(* IEC 61131-3 sources: volt/packages/volt-lsp-iec/test-corpus/lenze-mid/Device/Plc Logic/Application/Library Manager/CAA Device Diagnosis, 56 files *)

(* ---- BUS_INFO.dut ---- *)
TYPE BUS_INFO :
STRUCT
	ETYPE : BUS_TYPE;
	IDSYSTEM : CAA.IDENT;
	IDINSTANCE : CAA.IDENT;
END_STRUCT
END_TYPE

(* ---- BUS_STATE.dut ---- *)
TYPE BUS_STATE :
(
	UNKNOWN,
	STOPPED,
	RUNNING,
	ERROR,
	DISABLED
);
END_TYPE

(* ---- BUS_TYPE.dut ---- *)
TYPE BUS_TYPE :
(
	UNKNOWN := 16#0,
	PROFIBUS_DP := 16#1,
	CAN := 16#2,
	CANOPEN := 16#3,
	DEVICENET := 16#4,
	ETHERCAT := 16#5,
	PROFINET_IO := 16#6,
	ETHERNET_IP := 16#7,
	SERCOSII := 16#8,
	SERCOSIII := 16#9,
	MODBUS_TCP := 16#A,
	MODBUS_RTU := 16#B,
	AS_INTERFACE := 16#C,
	INTERBUS := 16#D,
	J1939 := 16#E,
	LON := 16#F,
	CC_LINK := 16#10,
	POWERLINK := 16#11,
	ETHERNET := 16#12,
	SERIAL_LINE := 16#13,
	VEN_SPEC := 16#14,
	FIRST_MF := 16#8000,
	LAST := 16#FFFF
);
END_TYPE

(* ---- DED_PNS_SUBMODULE_CFG.dut ---- *)
TYPE DED_PNS_SUBMODULE_CFG :
STRUCT
	UISLOT : UINT;
	UISUBSLOT : UINT;
	ULMODULEID : UDINT;
	ULSUBMODULEID : UDINT;
	ULPROVDATALEN : UDINT;
	ULCONSDATALEN : UDINT;
END_STRUCT
END_TYPE

(* ---- DEVICE_INFO.dut ---- *)
TYPE DEVICE_INFO :
STRUCT
	ETYPE : DEVICE_TYPE;
	IDSYSTEM : CAA.IDENT;
	IDINSTANCE : CAA.IDENT;
END_STRUCT
END_TYPE

(* ---- DEVICE_STATE.dut ---- *)
TYPE DEVICE_STATE :
(
	UNKNOWN,
	STOPPED,
	RUNNING,
	ERROR,
	DISABLED,
	NOT_CONFIGURED,
	CONFIGURED,
	NOT_FOUND
);
END_TYPE

(* ---- DEVICE_TRANSITION_STATE.dut ---- *)
TYPE DEVICE_TRANSITION_STATE :
(
	START,
	STOP,
	RESET
);
END_TYPE

(* ---- DEVICE_TYPE.dut ---- *)
TYPE DEVICE_TYPE :
(
	UNKNOWN := 16#0,
	FIELDBUS_MASTER := 16#1,
	FIELDBUS_SLAVE := 16#2,
	SAFETY_DEVICE := 16#3,
	SM_DEVICE := 16#4,
	SOFT_VISION_DEVICE := 16#5,
	DTM_DEVICE := 16#6,
	SPEC_IO_MODULE := 16#7,
	PLC := 16#1000,
	SAFETY_PLC := 16#1002,
	DRIVE := 16#1003,
	PARAM_DEVICE := 16#1004,
	HMI := 16#1005,
	SM_PLC := 16#1006
);
END_TYPE

(* ---- ERROR.dut ---- *)
TYPE ERROR :
(
	NO_ERROR := 0,
	FIRST_ERROR := 1300,
	TIME_OUT := 1301,
	ABORT := 1302,
	REF_INVALID := 1303,
	NOT_SUPPORTED := 1304,
	ERROR_IO := 1305,
	PARAM_INVALID := 1306,
	NODE_NOT_EXISTING := 1307,
	NO_MEMORY := 1308,
	ADR_NOT_FOUND := 1309,
	INST_NOT_FOUND := 1310,
	NO_DATA := 1311,
	OPERATION_INVALID := 1312,
	FIRST_MF := 1350,
	LAST_ERROR := 1399
);
END_TYPE

(* ---- ERROR_INFO.dut ---- *)
TYPE ERROR_INFO :
STRUCT
	IDERRORCODE : CAA.IDENT;
END_STRUCT
END_TYPE

(* ---- LOG_ENTRY.dut ---- *)
TYPE LOG_ENTRY :
STRUCT
	TKTIMESTAMP : CAA.TICK;
	IDMESSAGE : CAA.IDENT;
	IDSOURCE : CAA.IDENT;
END_STRUCT
END_TYPE

(* ---- LOGGER_MODE.dut ---- *)
TYPE LOGGER_MODE :
(
	LINEAR,
	CIRCULAR
);
END_TYPE

(* ---- PROC_CMD.dut ---- *)
TYPE PROC_CMD :
(
	NONE := 0,
	EXECUTE,
	ABORT
);
END_TYPE

(* ---- PROC_STATE.dut ---- *)
TYPE PROC_STATE :
(
	DORMAND := 0,
	BUSY,
	DONE,
	ABORTED,
	ERROR
);
END_TYPE

(* ---- QOS_INFO.dut ---- *)
TYPE QOS_INFO :
STRUCT
	CTERROR : CAA.COUNT;
	USIBUSLOAD : USINT;
END_STRUCT
END_TYPE

(* ---- TIDENTIFICATIONPARAMETER.dut ---- *)
TYPE TIDENTIFICATIONPARAMETER :
STRUCT
	IPADDRESS : ARRAY [0..3] OF BYTE;
	SUBNETMASK : ARRAY [0..3] OF BYTE;
	DEFAULTGATEWAY : ARRAY [0..3] OF BYTE;
	MACADDRESS : ARRAY [0..5] OF BYTE;
	STATIONNAME : STRING;
END_STRUCT
END_TYPE

(* ---- TISOCHRONEMODE.dut ---- *)
TYPE TISOCHRONEMODE :
STRUCT
	T_DC_BASE : UINT;
	T_DC_MIN : UINT;
	T_DC_MAX : UINT;
	T_IO_BASE : UDINT;
	T_IO_INPUTMIN : UDINT;
	T_IO_OUTPUTMIN : UDINT;
	ISOCHRONEMODEREQUIRED : BOOL;
END_STRUCT
END_TYPE

(* ---- TMODULEPARAMETER.dut ---- *)
TYPE TMODULEPARAMETER :
STRUCT
	MODULEIDENTNUMBER : UDINT;
	SLOTNUMBER : UINT;
	UINUMBERSUBMODULES : UINT;
END_STRUCT
END_TYPE

(* ---- TSLAVEPARAMETER.dut ---- *)
TYPE TSLAVEPARAMETER :
STRUCT
	UIDEVICEID : UINT;
	UIVENDORID : UINT;
	IDENTIFICATION : TIdentificationParameter;
	RTCLASS : UINT;
	VLANID : UINT;
	VLANPRIORITY : UINT;
	SENDCLOCK : UINT;
	REDUCTIONRATIO : UINT;
	WATCHDOGINTERVAL : UINT;
	MULTIPLEWRITESUPPORTED : BOOL;
	IOXSREQUIRED : BOOL;
	MAXINPUTLENGTH : UINT;
	MAXOUTPUTLENGTH : UINT;
	MAXDATALENGTH : UINT;
	UIMINSLAVEINTERVAL : UINT;
	UIOBJECTUUIDINSTANCE : UINT;
END_STRUCT
END_TYPE

(* ---- TVIRTUALSUBMODULE.dut ---- *)
TYPE TVIRTUALSUBMODULE :
STRUCT
	SUBMODULEIDENTNUMBER : UDINT;
	SUBSLOTNUMBER : UINT;
	API : UDINT;
	PROFISAFESUPPORTED : BOOL;
	ISOCHRONEMODE : TIsochroneMode;
	UINUMBERRDI : UINT;
	UISUBMODULEPROP : UINT;
	USIIOPSLEN : USINT;
	USIIOCSLEN : USINT;
END_STRUCT
END_TYPE

(* ---- DEVICEDIAGNOSISGLOBALS.gvl ---- *)
VAR_GLOBAL
	G_ITFROOTINODEINST : POINTER TO INode;
	G_ITFROOTNODECOUNT : UDINT;
END_VAR

(* ---- ERROR_CODES.gvl ---- *)
VAR_GLOBAL
	EC_NO_ERROR : CAA.IDENT := 16#0;
	EC_FIRST_INFO : CAA.IDENT := 16#1000;
	EC_LAST_INFO : CAA.IDENT := 16#1FFF;
	EC_FIRST_WARNING : CAA.IDENT := 16#2000;
	EC_LAST_WARNING : CAA.IDENT := 16#2FFF;
	EC_FIRST_ERROR : CAA.IDENT := 16#3000;
	EC_LAST_ERROR : CAA.IDENT := 16#3FFF;
	EC_FIRST_EMCY : CAA.IDENT := 16#4000;
	EC_LAST_EMCY : CAA.IDENT := 16#4FFF;
END_VAR

(* ---- VERSIONCONSTANTS.gvl ---- *)
VAR_GLOBAL
	GC_BYVERSION : BYTE := 1;
	GC_BYVERSION_1 : BYTE := 1;
END_VAR

(* ---- IBUS.itf ---- *)
INTERFACE IBUS
END_INTERFACE

METHOD GETBUSDIAGNOSISINFO : ERROR
VAR_INPUT
	PDATA : CAA.PVOID;
	SZSIZE : CAA.SIZE;
END_VAR
VAR_OUTPUT
	SZCOUNT : CAA.SIZE;
END_VAR
END_METHOD

METHOD GETBUSERRORASYNC : PROC_STATE
VAR_INPUT
	ECMD : PROC_CMD;
END_VAR
VAR_OUTPUT
	EERROR : ERROR;
END_VAR
VAR_IN_OUT
	ERIBUSERROR : ERROR_INFO;
END_VAR
END_METHOD

METHOD GETBUSINFO : ERROR
VAR_IN_OUT
	BUIINFO : BUS_INFO;
END_VAR
END_METHOD

METHOD GETBUSSTATE : BUS_STATE
VAR_OUTPUT
	XDIAGNOSISINFOAVAILABLE : BOOL;
	EERROR : ERROR;
END_VAR
END_METHOD

METHOD GETQOS : ERROR
VAR_IN_OUT
	QUALITYINFO : QOS_INFO;
END_VAR
END_METHOD

METHOD GETSPECIFICBUSSTATE : ERROR
VAR_INPUT
	PDATA : CAA.PVOID;
	SZSIZE : CAA.SIZE;
END_VAR
VAR_OUTPUT
	SZCOUNT : CAA.SIZE;
END_VAR
END_METHOD

(* ---- IDEVICE.itf ---- *)
INTERFACE IDEVICE
END_INTERFACE

METHOD GETDEVICEDIAGNOSISINFO : ERROR
VAR_INPUT
	PDATA : CAA.PVOID;
	SZSIZE : CAA.SIZE;
END_VAR
VAR_OUTPUT
	SZCOUNT : CAA.SIZE;
END_VAR
END_METHOD

METHOD GETDEVICEERRORASYNC : PROC_STATE
VAR_INPUT
	ECMD : PROC_CMD;
END_VAR
VAR_OUTPUT
	EERROR : ERROR;
END_VAR
VAR_IN_OUT
	ERIDEVICEERROR : ERROR_INFO;
END_VAR
END_METHOD

METHOD GETDEVICEINFO : ERROR
VAR_IN_OUT
	DEIINFO : DEVICE_INFO;
END_VAR
END_METHOD

METHOD GETDEVICESTATE : DEVICE_STATE
VAR_OUTPUT
	XDIAGNOSISINFOAVAILABLE : BOOL;
	EERROR : ERROR;
END_VAR
END_METHOD

METHOD SETCOMMUNICATIONSTATE : ERROR
VAR_INPUT
	EREQUESTEDSTATE : DEVICE_TRANSITION_STATE;
END_VAR
END_METHOD

METHOD GETSPECIFICDEVICEERRORASYNC : PROC_STATE
VAR_INPUT
	ECMD : PROC_CMD;
	PDATA : CAA.PVOID;
	SZSIZE : CAA.SIZE;
END_VAR
VAR_OUTPUT
	SZCOUNT : CAA.SIZE;
	EERROR : ERROR;
END_VAR
END_METHOD

METHOD GETSPECIFICDEVICESTATE : ERROR
VAR_INPUT
	PDATA : CAA.PVOID;
	SZSIZE : CAA.SIZE;
END_VAR
VAR_OUTPUT
	SZCOUNT : CAA.SIZE;
END_VAR
END_METHOD

(* ---- IDEVICE2.itf ---- *)
INTERFACE IDEVICE2
END_INTERFACE

METHOD CHECKCURRENTSUPPORTEDCOMMUNICATIONSTATE : BOOL
VAR_INPUT
	EREQUESTEDSTATE : DEVICE_TRANSITION_STATE;
END_VAR
END_METHOD

METHOD CHECKSUPPORTEDCOMMUNICATIONSTATE : BOOL
VAR_INPUT
	EREQUESTEDSTATE : DEVICE_TRANSITION_STATE;
END_VAR
END_METHOD

(* ---- ILOGGER.itf ---- *)
INTERFACE ILOGGER
END_INTERFACE

METHOD DISABLELOGGER : ERROR
END_METHOD

METHOD ENABLELOGGER : ERROR
VAR_INPUT
	EMODE : LOGGER_MODE;
	CTMAXLOGMESSAGES : CAA.COUNT;
END_VAR
END_METHOD

METHOD GETLOGENTRY : ERROR
VAR_IN_OUT
	LOGENTRY : LOG_ENTRY;
END_VAR
END_METHOD

(* ---- INODE.itf ---- *)
INTERFACE INODE
END_INTERFACE

METHOD GETCHILD : INode
VAR_INPUT
	UDIINDEX : UDINT;
END_VAR
END_METHOD

METHOD INITIALIZE_DIAG : UDINT
VAR_INPUT
	PCONNECTOR : POINTER TO IoConfigConnector;
	NCONNECTORCOUNT : DINT;
	PARENT : POINTER TO INode;
	CHILDREN : POINTER TO INode;
	UDICHILDCOUNT : UDINT;
END_VAR
END_METHOD

(* ---- IRECONFIGUREPROVIDER.itf ---- *)
INTERFACE IRECONFIGUREPROVIDER
END_INTERFACE

METHOD RECONFIGUREASYNC : PROC_STATE
VAR_INPUT
	ECMD : PROC_CMD;
	ITFSENDER : INode;
END_VAR
VAR_OUTPUT
	EERROR : ERROR;
END_VAR
END_METHOD

METHOD REGISTERIRPCHILD : ERROR
VAR_INPUT
	ITFCHILD : IReconfigureProvider;
END_VAR
END_METHOD

(* ---- ISTACK.itf ---- *)
INTERFACE ISTACK
END_INTERFACE

METHOD GETBUSSCANASYNC : PROC_STATE
VAR_INPUT
	ECMD : PROC_CMD;
END_VAR
VAR_OUTPUT
	ITFFIRSTDEVICE : INode;
	EERROR : ERROR;
END_VAR
END_METHOD

METHOD GETLOGGER : ILogger
VAR_OUTPUT
	EERROR : ERROR;
END_VAR
END_METHOD

(* ---- CANRECONFIGURE.pou ---- *)
FUNCTION CANRECONFIGURE : BOOL
VAR_INPUT
	ITFNODE : INode;
END_VAR
END_FUNCTION

(* ---- GETDEVICENAMESTRING.pou ---- *)
FUNCTION GETDEVICENAMESTRING : STRING
VAR_INPUT
	ITFNODE : INode;
END_VAR
END_FUNCTION

(* ---- GETDEVICENAMEWSTRING.pou ---- *)
FUNCTION GETDEVICENAMEWSTRING : WSTRING
VAR_INPUT
	ITFNODE : INode;
END_VAR
END_FUNCTION

(* ---- GETNEXTNODE.pou ---- *)
FUNCTION GETNEXTNODE : INode
VAR_INPUT
	ITFCURRENT : INode;
END_VAR
END_FUNCTION

(* ---- GETNODEDEPTH.pou ---- *)
FUNCTION GETNODEDEPTH : INT
VAR_INPUT
	ITFNODE : INode;
END_VAR
END_FUNCTION

(* ---- GETROOT.pou ---- *)
FUNCTION GETROOT : INode
END_FUNCTION

(* ---- GETSUPPLIERVERSION.pou ---- *)
FUNCTION GETSUPPLIERVERSION : WORD
VAR_INPUT
	XDUMMY : BOOL;
END_VAR
END_FUNCTION

(* ---- INODE_TO_IBUS.pou ---- *)
FUNCTION INODE_TO_IBUS : IBus
VAR_INPUT
	ITFNODE : INode;
END_VAR
END_FUNCTION

(* ---- INODE_TO_IDEVICE.pou ---- *)
FUNCTION INODE_TO_IDEVICE : IDevice
VAR_INPUT
	ITFNODE : INode;
END_VAR
END_FUNCTION

(* ---- INODE_TO_IDEVICE2.pou ---- *)
FUNCTION INODE_TO_IDEVICE2 : IDevice2
VAR_INPUT
	ITFNODE : INode;
END_VAR
END_FUNCTION

(* ---- INODE_TO_ISTACK.pou ---- *)
FUNCTION INODE_TO_ISTACK : IStack
VAR_INPUT
	ITFNODE : INode;
END_VAR
END_FUNCTION

(* ---- ISCONNECTORENABLED.pou ---- *)
FUNCTION ISCONNECTORENABLED : BOOL
VAR_INPUT
	PCONNECTOR : POINTER TO IoStandard.IoConfigConnector;
END_VAR
END_FUNCTION

(* ---- CAADIAGDEVICEDEFAULT.pou ---- *)
FUNCTION_BLOCK CAADIAGDEVICEDEFAULT EXTENDS CAADiagTreeBase
VAR
	M_DIAG : CAADiagnosisBase;
	_DEIINFO : DEVICE_INFO;
END_VAR
END_FUNCTION_BLOCK

METHOD CHECKCURRENTSUPPORTEDCOMMUNICATIONSTATE : BOOL
VAR_INPUT
	EREQUESTEDSTATE : DEVICE_TRANSITION_STATE;
END_VAR
END_METHOD

METHOD CHECKSUPPORTEDCOMMUNICATIONSTATE : BOOL
VAR_INPUT
	EREQUESTEDSTATE : DEVICE_TRANSITION_STATE;
END_VAR
END_METHOD

METHOD GETDEVICEDIAGNOSISINFO : ERROR
VAR_INPUT
	PDATA : CAA.PVOID;
	SZSIZE : CAA.SIZE;
END_VAR
VAR_OUTPUT
	SZCOUNT : CAA.SIZE;
END_VAR
END_METHOD

METHOD GETDEVICEERRORASYNC : PROC_STATE
VAR_INPUT
	ECMD : PROC_CMD;
END_VAR
VAR_OUTPUT
	EERROR : ERROR;
END_VAR
VAR_IN_OUT
	ERIDEVICEERROR : ERROR_INFO;
END_VAR
END_METHOD

METHOD GETDEVICEINFO : ERROR
VAR_IN_OUT
	DEIINFO : DEVICE_INFO;
END_VAR
END_METHOD

METHOD GETDEVICESTATE : DEVICE_STATE
VAR_OUTPUT
	XDIAGNOSISINFOAVAILABLE : BOOL;
	EERROR : ERROR;
END_VAR
END_METHOD

METHOD GETPROFINETDEVICEINFO : ERROR
VAR_IN_OUT
	DEIINFO : DEVICE_INFO;
END_VAR
END_METHOD

METHOD GETSPECIFICDEVICEERRORASYNC : PROC_STATE
VAR_INPUT
	ECMD : PROC_CMD;
	PDATA : CAA.PVOID;
	SZSIZE : CAA.SIZE;
END_VAR
VAR_OUTPUT
	SZCOUNT : CAA.SIZE;
	EERROR : ERROR;
END_VAR
END_METHOD

METHOD GETSPECIFICDEVICESTATE : ERROR
VAR_INPUT
	PDATA : CAA.PVOID;
	SZSIZE : CAA.SIZE;
END_VAR
VAR_OUTPUT
	SZCOUNT : CAA.SIZE;
END_VAR
END_METHOD

METHOD INITIALIZE_DIAG : UDINT
VAR_INPUT
	PCONNECTOR : POINTER TO IoConfigConnector;
	NCONNECTORCOUNT : DINT;
	PARENT : POINTER TO INode;
	CHILDREN : POINTER TO INode;
	UDICHILDCOUNT : UDINT;
END_VAR
END_METHOD

METHOD SETCOMMUNICATIONSTATE : ERROR
VAR_INPUT
	EREQUESTEDSTATE : DEVICE_TRANSITION_STATE;
END_VAR
END_METHOD

(* ---- CAADIAGNOSISBASE.pou ---- *)
FUNCTION_BLOCK CAADIAGNOSISBASE
VAR
	M_NCOUNT : DINT;
	M_PCONNECTOR : POINTER TO IoConfigConnector;
	BUSLOGGER : Logger;
END_VAR
END_FUNCTION_BLOCK

METHOD CALCIPADRUDINT : UDINT
VAR_INPUT
	PABY : POINTER TO ARRAY [0..3] OF BYTE;
END_VAR
END_METHOD

METHOD GETBUSINFO : ERROR
VAR_IN_OUT
	BUIINFO : BUS_INFO;
END_VAR
END_METHOD

METHOD GETBUSSCANASYNC : PROC_STATE
VAR_INPUT
	ECMD : PROC_CMD;
END_VAR
VAR_OUTPUT
	ITFFIRSTDEVICE : INode;
	EERROR : ERROR;
END_VAR
END_METHOD

METHOD GETBUSSTATE : BUS_STATE
VAR_OUTPUT
	XDIAGNOSISINFOAVAILABLE : BOOL;
	EERROR : ERROR;
END_VAR
END_METHOD

METHOD GETDEVICEINFO : ERROR
VAR_IN_OUT
	DEIINFO : DEVICE_INFO;
END_VAR
END_METHOD

METHOD GETERRORASYNC : PROC_STATE
VAR_INPUT
	ECMD : PROC_CMD;
END_VAR
VAR_OUTPUT
	EERROR : ERROR;
END_VAR
VAR_IN_OUT
	ERIERROR : ERROR_INFO;
END_VAR
END_METHOD

METHOD GETSPECIFICDEVICEERRORASYNC : PROC_STATE
VAR_INPUT
	ECMD : PROC_CMD;
	PDATA : CAA.PVOID;
	SZSIZE : CAA.SIZE;
END_VAR
VAR_OUTPUT
	SZCOUNT : CAA.SIZE;
	EERROR : ERROR;
END_VAR
END_METHOD

METHOD GETSTATE : DEVICE_STATE
VAR_OUTPUT
	XDIAGNOSISINFOAVAILABLE : BOOL;
	EERROR : ERROR;
END_VAR
END_METHOD

METHOD INITIALIZE_DIAG : UDINT
VAR_INPUT
	PCONNECTOR : POINTER TO IoConfigConnector;
	NCOUNT : DINT;
END_VAR
END_METHOD

(* ---- CAADIAGTREEBASE.pou ---- *)
FUNCTION_BLOCK CAADIAGTREEBASE
VAR
	M_PARENT : POINTER TO INode := CAA.gc_pNULL;
	M_CHILDREN : POINTER TO INode := CAA.gc_pNULL;
	M_UDICHILDCOUNT : UDINT;
	M_UDICHILDINDEX : UDINT;
	M_NCOUNT : DINT;
	M_PCONNECTOR : POINTER TO IoConfigConnector;
	CHILDNODECOUNT : CAA.Count;
	CONNECTOR : POINTER TO IoConfigConnector;
	ENABLE : BOOL;
	FIRSTCHILDNODE : INode;
	INDEX : UDINT;
	ISROOTNODE : BOOL;
	NEXTSIBLINGNODE : INode;
	PARENTNODE : INode;
	SIBLINGNODECOUNT : CAA.Count;
END_VAR
END_FUNCTION_BLOCK

METHOD GETCHILD : INode
VAR_INPUT
	UDIINDEX : UDINT;
END_VAR
END_METHOD

METHOD INITIALIZE_DIAG : UDINT
VAR_INPUT
	PCONNECTOR : POINTER TO IoConfigConnector;
	NCONNECTORCOUNT : DINT;
	PARENT : POINTER TO INode;
	CHILDREN : POINTER TO INode;
	UDICHILDCOUNT : UDINT;
END_VAR
END_METHOD

(* ---- CAARECONFIGUREBASE.pou ---- *)
FUNCTION_BLOCK CAARECONFIGUREBASE
VAR
	_ITFMYNODE : INode;
	_ITFSIBLING : IReconfigureProvider;
	_ITFFIRSTCHILDIRP : IReconfigureProvider;
	_BYRECONFIGURESTATE : BYTE;
	_XRECONFIGUREERROR : BOOL;
	_BYRECONFIGURECHILDRENSTATE : BYTE;
	_XRECONFIGURECHILDRENERROR : BOOL;
	_BYRECONFIGUREIODRIVERSTATE : BYTE;
	_UDIIOMGRASYNCSTATE : UDINT := CmpAsyncMgr.ASYNCSTATE_PENDING;
	_UDIBEGINCOUNT : UDINT;
	RECONFIGUREACTIVE : BOOL;
	SIBLINGIRP : IReconfigureProvider;
END_VAR
END_FUNCTION_BLOCK

METHOD BEGINRECONFIGURE
VAR_INPUT
	ITFSENDER : INode;
END_VAR
END_METHOD

METHOD ENDRECONFIGURE
VAR_INPUT
	ITFSENDER : INode;
END_VAR
END_METHOD

METHOD INITIALIZE_DIAG : ERROR
VAR_INPUT
	ITFNODE : INode;
END_VAR
END_METHOD

METHOD UPDATEENABLEFLAGS
END_METHOD

METHOD RECONFIGUREASYNC : PROC_STATE
VAR_INPUT
	ECMD : PROC_CMD;
	ITFSENDER : INode;
END_VAR
VAR_OUTPUT
	EERROR : ERROR;
END_VAR
END_METHOD

METHOD REGISTERIRPCHILD : ERROR
VAR_INPUT
	ITFCHILD : IReconfigureProvider;
END_VAR
END_METHOD

METHOD RECONFIGURECHILDRENASYNC : PROC_STATE
VAR_INPUT
	ECMD : PROC_CMD;
	ITFSENDER : INode;
END_VAR
VAR_OUTPUT
	EERROR : ERROR;
END_VAR
END_METHOD

METHOD RECONFIGUREIODRIVERASYNC : PROC_STATE
VAR_INPUT
	ECMD : PROC_CMD;
	ITFSENDER : INode;
END_VAR
VAR_OUTPUT
	EERROR : ERROR;
END_VAR
END_METHOD

(* ---- ETRIG.pou ---- *)
FUNCTION_BLOCK ETRIG
VAR_INPUT
	XEXECUTE : BOOL;
END_VAR
VAR_OUTPUT
	XDONE : BOOL;
	XBUSY : BOOL;
	XERROR : BOOL;
END_VAR
VAR
	XPREVIOUSEXECUTE : BOOL;
	XPREVIOUSABORTINPROGRESS : BOOL;
	XABORTINPROGRESS : BOOL;
	IERROR : INT;
END_VAR
END_FUNCTION_BLOCK

METHOD PRVABORT : BOOL
END_METHOD

METHOD PRVCYCLICACTION : BOOL
END_METHOD

METHOD PRVRESETOUTPUTS : BOOL
END_METHOD

METHOD PRVSTART : BOOL
END_METHOD

(* ---- ETRIGA.pou ---- *)
FUNCTION_BLOCK ETRIGA
VAR_INPUT
	XEXECUTE : BOOL;
	XABORT : BOOL;
END_VAR
VAR_OUTPUT
	XDONE : BOOL;
	XBUSY : BOOL;
	XERROR : BOOL;
	XABORTED : BOOL;
END_VAR
VAR
	XPREVIOUSABORTINPROGRESS : BOOL;
	XPREVIOUSEXECUTE : BOOL;
	XABORTINPROGRESS : BOOL;
	IERROR : INT;
END_VAR
END_FUNCTION_BLOCK

METHOD PRVABORT : BOOL
END_METHOD

METHOD PRVCYCLICACTION : BOOL
END_METHOD

METHOD PRVRESETOUTPUTS : BOOL
END_METHOD

METHOD PRVSTART : BOOL
END_METHOD

(* ---- GETBUSERROR.pou ---- *)
FUNCTION_BLOCK GETBUSERROR EXTENDS ETrigA
VAR_INPUT
	ITFNODE : INode;
END_VAR
VAR_OUTPUT
	EERROR : ERROR;
	EINBUSERROR : ERROR_INFO;
END_VAR
VAR
	ITFBUS : IBus;
END_VAR
END_FUNCTION_BLOCK

METHOD PRVABORT : BOOL
END_METHOD

METHOD PRVCYCLICACTION : BOOL
END_METHOD

METHOD PRVRESETOUTPUTS : BOOL
END_METHOD

METHOD PRVSTART : BOOL
END_METHOD

(* ---- GETBUSSCAN.pou ---- *)
FUNCTION_BLOCK GETBUSSCAN EXTENDS ETrigA
VAR_INPUT
	ITFNODE : INode;
END_VAR
VAR_OUTPUT
	EERROR : ERROR;
	ITFFIRSTDEVICE : INode;
END_VAR
VAR
	_ITFSTACK : IStack;
END_VAR
END_FUNCTION_BLOCK

METHOD PRVABORT : BOOL
END_METHOD

METHOD PRVCYCLICACTION : BOOL
END_METHOD

METHOD PRVRESETOUTPUTS : BOOL
END_METHOD

METHOD PRVSTART : BOOL
END_METHOD

(* ---- GETDEVICEERROR.pou ---- *)
FUNCTION_BLOCK GETDEVICEERROR EXTENDS ETrigA
VAR_INPUT
	ITFNODE : INode;
END_VAR
VAR_OUTPUT
	EERROR : ERROR;
	EINDEVICEERROR : ERROR_INFO;
END_VAR
VAR
	ITFDEVICE : IDevice;
END_VAR
END_FUNCTION_BLOCK

METHOD PRVABORT : BOOL
END_METHOD

METHOD PRVCYCLICACTION : BOOL
END_METHOD

METHOD PRVRESETOUTPUTS : BOOL
END_METHOD

METHOD PRVSTART : BOOL
END_METHOD

(* ---- GETIDEVICEINSTBYIOADDR.pou ---- *)
FUNCTION_BLOCK GETIDEVICEINSTBYIOADDR EXTENDS ETrigA
VAR_INPUT
	DWADDRESS : DWORD;
	DWBITOFFSET : DWORD;
END_VAR
VAR_OUTPUT
	ITFDEVICE : IDevice;
END_VAR
VAR
	M_PCONNECTOR : POINTER TO IoConfigConnector;
	M_PTASKMAPLIST : POINTER TO IoConfigTaskMap;
	M_NTASKMAPLISTCOUNT : DINT;
	M_ISTATE : INT;
	M_HCALLBACK : SysTypes.RTS_IEC_HANDLE := SysTypes.RTS_INVALID_HANDLE;
END_VAR
END_FUNCTION_BLOCK

METHOD EVENTCALLBACK : UDINT
VAR_INPUT
	PEVENTPARAM : POINTER TO EventParam;
END_VAR
END_METHOD

METHOD FB_EXIT : BOOL
VAR_INPUT
	BINCOPYCODE : BOOL;
END_VAR
END_METHOD

METHOD FB_INIT : BOOL
VAR_INPUT
	BINITRETAINS : BOOL;
	BINCOPYCODE : BOOL;
END_VAR
END_METHOD

METHOD PRVABORT : BOOL
END_METHOD

METHOD PRVCYCLICACTION : BOOL
END_METHOD

METHOD PRVRESETOUTPUTS : BOOL
END_METHOD

METHOD PRVSTART : BOOL
END_METHOD

(* ---- GETSPECIFICDEVICEERROR.pou ---- *)
FUNCTION_BLOCK GETSPECIFICDEVICEERROR EXTENDS ETrigA
VAR_INPUT
	ITFNODE : INode;
	PDATA : CAA.PVOID;
END_VAR
VAR_OUTPUT
	EERROR : ERROR;
END_VAR
VAR_IN_OUT
	SZSIZE : CAA.SIZE;
END_VAR
VAR
	ITFDEVICE : IDevice;
END_VAR
END_FUNCTION_BLOCK

METHOD PRVABORT : BOOL
END_METHOD

METHOD PRVCYCLICACTION : BOOL
END_METHOD

METHOD PRVRESETOUTPUTS : BOOL
END_METHOD

METHOD PRVSTART : BOOL
END_METHOD

(* ---- LOGGER.pou ---- *)
FUNCTION_BLOCK LOGGER
END_FUNCTION_BLOCK

METHOD DISABLELOGGER : ERROR
END_METHOD

METHOD ENABLELOGGER : ERROR
VAR_INPUT
	EMODE : LOGGER_MODE;
	CTMAXLOGMESSAGES : CAA.COUNT;
END_VAR
END_METHOD

METHOD GETLOGENTRY : ERROR
VAR_IN_OUT
	LOGENTRY : LOG_ENTRY;
END_VAR
END_METHOD

(* ---- RECONFIGURE.pou ---- *)
FUNCTION_BLOCK RECONFIGURE EXTENDS ETrig
VAR_INPUT
	ITFNODE : INode;
END_VAR
VAR_OUTPUT
	EERROR : ERROR;
END_VAR
VAR
	_ITFRECONFIGURE : IReconfigureProvider;
END_VAR
END_FUNCTION_BLOCK

METHOD PRVABORT : BOOL
END_METHOD

METHOD PRVCYCLICACTION : BOOL
END_METHOD

METHOD PRVRESETOUTPUTS : BOOL
END_METHOD

METHOD PRVSTART : BOOL
END_METHOD

(* ---- RECURSIVEHELPER.pou ---- *)
FUNCTION_BLOCK RECURSIVEHELPER
END_FUNCTION_BLOCK

METHOD UPDATEENABLEFLAGSRECURSIVE
VAR_INPUT
	ITFNODE : INode;
	XPARENTENABLE : BOOL;
END_VAR
END_METHOD
